(* IEC 61131-3 sources: POMIRTS_lab3/AS/Library/ETHERNET, 3 files *)

(* ---- ETHERNET.typ ---- *)
(********************************************************************
 * COPYRIGHT (C) BERNECKER + RAINER, AUSTRIA, A-5142 EGGELSBERG
 ********************************************************************
 * Library: Ethernet
 * File: Ethernet.typ
 * Created: 11.11.2003
 ********************************************************************
 * Global data types of library Ethernet
 ********************************************************************)
TYPE
	ETHattachment_typ : STRUCT
		type	: USINT ;
		len	: UDINT ;
		pName	: UDINT ;
		pData	: UDINT ;
	END_STRUCT;
	ETHstatSG3_typ : STRUCT
		l_int	: UDINT ;
		l_rint	: UDINT ;
		l_tint	: UDINT ;
		l_babl	: UINT ;
		l_cerr	: UINT ;
		l_miss	: UINT ;
		l_memr	: UINT ;
		r_fram	: UINT ;
		r_oflo	: UINT ;
		r_crc	: UINT ;
		r_buff	: UINT ;
		t_buff	: UINT ;
		t_uflo	: UINT ;
		t_lcol	: UINT ;
		t_lcar	: UINT ;
		t_rtry	: UINT ;
		ni_anno	: UINT ;
		ni_init	: UINT ;
		ni_send	: UINT ;
		ni_getp	: UINT ;
		ni_retp	: UINT ;
		ni_bcst	: UINT ;
		ni_poll	: UINT ;
		irq_mean	: UINT ;
		irq_min	: UINT ;
		irq_max	: UINT ;
		irq_t1	: UINT ;
		irq_timena	: UINT ;
		errgtnobuf	: UINT ;
		err_1_1	: UINT ;
		err_1_2	: UINT ;
		err_1_3	: UINT ;
		errxmtnull	: UINT ;
		errsndown	: UINT ;
		errsndsize	: UINT ;
		lancerrnobuf	: UINT ;
		lanceinit	: UINT ;
		terr	: UINT ;
		ni_gtbuf	: UINT ;
		brcast_cnt	: UINT ;
		brcastmax_cnt	: UINT ;
		brcast_stop	: UINT ;
		brcast_tick	: UINT ;
	END_STRUCT;
	ETHstatSG4_typ : STRUCT
		p_recv	: UDINT ;
		e_recv	: UDINT ;
		p_send	: UDINT ;
		e_send	: UDINT ;
		collisions	: UDINT ;
		b_recv	: UDINT ;
		b_send	: UDINT ;
		p_recv_mc	: UDINT ;
		p_send_mc	: UDINT ;
		iqdrops	: UDINT ;
		noproto	: UDINT ;
		lastchange	: UDINT ;
	END_STRUCT;
	TCPQ_dcmd_typ : STRUCT
		response	: UINT ;
		error	: UDINT ;
		buffer	: UDINT ;
		buflng	: UDINT ;
		ipaddr	: UDINT ;
		socket	: UDINT ;
		port	: UINT ;
		wreserve	: UINT ;
		reserve	: ARRAY[0..7] OF UDINT ;
	END_STRUCT;
END_TYPE

(* ---- ETHERNET.fun ---- *)
(********************************************************************
 * COPYRIGHT (C) BERNECKER + RAINER, AUSTRIA, A-5142 EGGELSBERG
 ********************************************************************
 * Library: Ethernet
 * File: Ethernet.fun
 * Created: 11.11.2003
 ********************************************************************
 * Functions and function blocks of library Ethernet
 ********************************************************************)
FUNCTION_BLOCK ETHinfo
	VAR_INPUT
		enable	:BOOL;
	END_VAR
	VAR_OUTPUT
		statadr	:UDINT;
		ethadr	:UDINT;
		status	:UINT;
	END_VAR
END_FUNCTION_BLOCK
FUNCTION_BLOCK SMTPxsendmail
	VAR_INPUT
		enable	:BOOL;
		pReceiver	:UDINT;
		pSender	:UDINT;
		pIpaddr	:UDINT;
		pSubject	:UDINT;
		pText	:UDINT;
		pAttachment	:UDINT;
		AttachmentCount	:USINT;
		timeout	:UINT;
	END_VAR
	VAR_OUTPUT
		status	:UINT;
	END_VAR
	VAR
		pna_ok	:BOOL;
		state	:UINT;
		tickcount	:UDINT;
		initcount	:UDINT;
		dcmd	:TCPQ_dcmd_typ;
	END_VAR
END_FUNCTION_BLOCK
FUNCTION_BLOCK ETHxinfo
	VAR_INPUT
		enable	:BOOL;
		pDevice	:UDINT;
	END_VAR
	VAR_OUTPUT
		statadr	:UDINT;
		ethadr	:UDINT;
		status	:UINT;
	END_VAR
	VAR
		mac	:ARRAY[0..5] OF USINT;
	END_VAR
END_FUNCTION_BLOCK
FUNCTION_BLOCK TCPclose
	VAR_INPUT
		enable	:BOOL;
		cident	:UDINT;
	END_VAR
	VAR_OUTPUT
		status	:UINT;
	END_VAR
	VAR
		pna_ok	:BOOL;
		state	:UINT;
		tickcount	:UDINT;
		initcount	:UDINT;
		dcmd	:TCPQ_dcmd_typ;
	END_VAR
END_FUNCTION_BLOCK
FUNCTION_BLOCK TCPrecv
	VAR_INPUT
		enable	:BOOL;
		cident	:UDINT;
		buffer	:UDINT;
		mxbuflng	:UDINT;
	END_VAR
	VAR_OUTPUT
		status	:UINT;
		rxbuflng	:UDINT;
	END_VAR
	VAR
		pna_ok	:BOOL;
		state	:UINT;
		tickcount	:UDINT;
		initcount	:UDINT;
		dcmd	:TCPQ_dcmd_typ;
	END_VAR
END_FUNCTION_BLOCK
FUNCTION_BLOCK TCPsend
	VAR_INPUT
		enable	:BOOL;
		cident	:UDINT;
		buffer	:UDINT;
		buflng	:UDINT;
	END_VAR
	VAR_OUTPUT
		status	:UINT;
	END_VAR
	VAR
		pna_ok	:BOOL;
		state	:UINT;
		tickcount	:UDINT;
		initcount	:UDINT;
		dcmd	:TCPQ_dcmd_typ;
	END_VAR
END_FUNCTION_BLOCK
FUNCTION_BLOCK TCPclient
	VAR_INPUT
		enable	:BOOL;
		porta	:UINT;
		ipaddr	:UDINT;
		portb	:UINT;
	END_VAR
	VAR_OUTPUT
		status	:UINT;
		cident	:UDINT;
	END_VAR
	VAR
		pna_ok	:BOOL;
		state	:UINT;
		tickcount	:UDINT;
		initcount	:UDINT;
		dcmd	:TCPQ_dcmd_typ;
	END_VAR
END_FUNCTION_BLOCK
FUNCTION_BLOCK TCPserv
	VAR_INPUT
		enable	:BOOL;
		porta	:UINT;
	END_VAR
	VAR_OUTPUT
		status	:UINT;
		ipaddr	:UDINT;
		portb	:UINT;
		cident	:UDINT;
	END_VAR
	VAR
		pna_ok	:BOOL;
		state	:UINT;
		tickcount	:UDINT;
		initcount	:UDINT;
		dcmd	:TCPQ_dcmd_typ;
	END_VAR
END_FUNCTION_BLOCK
FUNCTION_BLOCK ICMPping
	VAR_INPUT
		enable	:BOOL;
		ipaddr	:UDINT;
		timeout	:UINT;
	END_VAR
	VAR_OUTPUT
		status	:UINT;
	END_VAR
	VAR
		pna_ok	:BOOL;
		state	:UINT;
		tickcount	:UDINT;
		initcount	:UDINT;
		dcmd	:TCPQ_dcmd_typ;
	END_VAR
END_FUNCTION_BLOCK
FUNCTION_BLOCK SMTPsendmail
	VAR_INPUT
		enable	:BOOL;
		pReceiver	:UDINT;
		pSender	:UDINT;
		pIpaddr	:UDINT;
		pSubject	:UDINT;
		pText	:UDINT;
		timeout	:UINT;
	END_VAR
	VAR_OUTPUT
		status	:UINT;
	END_VAR
	VAR
		pna_ok	:BOOL;
		state	:UINT;
		tickcount	:UDINT;
		initcount	:UDINT;
		dcmd	:TCPQ_dcmd_typ;
	END_VAR
END_FUNCTION_BLOCK
FUNCTION_BLOCK UDPclose
	VAR_INPUT
		enable	:BOOL;
		cident	:UDINT;
	END_VAR
	VAR_OUTPUT
		status	:UINT;
	END_VAR
	VAR
		pna_ok	:BOOL;
		state	:UINT;
		tickcount	:UDINT;
		initcount	:UDINT;
		dcmd	:TCPQ_dcmd_typ;
	END_VAR
END_FUNCTION_BLOCK
FUNCTION_BLOCK UDPopen
	VAR_INPUT
		enable	:BOOL;
		port	:UINT;
		pvpolladr	:UDINT;
	END_VAR
	VAR_OUTPUT
		status	:UINT;
		cident	:UDINT;
	END_VAR
	VAR
		pna_ok	:BOOL;
		state	:UINT;
		tickcount	:UDINT;
		initcount	:UDINT;
		dcmd	:TCPQ_dcmd_typ;
	END_VAR
END_FUNCTION_BLOCK
FUNCTION_BLOCK UDPrecv
	VAR_INPUT
		enable	:BOOL;
		cident	:UDINT;
		buffer	:UDINT;
		buflng	:UINT;
	END_VAR
	VAR_OUTPUT
		status	:UINT;
		ipaddr	:UDINT;
		rxbuflng	:UINT;
		port	:UINT;
	END_VAR
	VAR
		pna_ok	:BOOL;
		state	:UINT;
		tickcount	:UDINT;
		initcount	:UDINT;
		dcmd	:TCPQ_dcmd_typ;
	END_VAR
END_FUNCTION_BLOCK
FUNCTION_BLOCK UDPsend
	VAR_INPUT
		enable	:BOOL;
		cident	:UDINT;
		ipaddr	:UDINT;
		buffer	:UDINT;
		buflng	:UINT;
		port	:UINT;
	END_VAR
	VAR_OUTPUT
		status	:UINT;
	END_VAR
	VAR
		pna_ok	:BOOL;
		state	:UINT;
		tickcount	:UDINT;
		initcount	:UDINT;
		dcmd	:TCPQ_dcmd_typ;
	END_VAR
END_FUNCTION_BLOCK
FUNCTION_BLOCK ETHnode
	VAR_INPUT
		enable	:BOOL;
	END_VAR
	VAR_OUTPUT
		status	:UINT;
		nodenr	:USINT;
		ipaddr	:UDINT;
	END_VAR
	VAR
		address1	:UDINT;
		address2	:UDINT;
	END_VAR
END_FUNCTION_BLOCK

(* ---- ETHERNET.var ---- *)
(********************************************************************
 * COPYRIGHT (C) BERNECKER + RAINER, AUSTRIA, A-5142 EGGELSBERG
 ********************************************************************
 * Library: Ethernet
 * File: Ethernet.var
 * Created: 11.11.2003
 ********************************************************************
 * Constants of library Ethernet
 ********************************************************************)
VAR CONSTANT
	ERR_ETH_SMTP_UNEXPECTED_RESPONSE	: UINT	:= 27232;
	ERR_ETH_SMTP_SERVER_NOTAVAILABLE	: UINT	:= 27230;
	ERR_ETH_SMTP_RECEIVER_NOT_ACCEPT	: UINT	:= 27234;
	ERR_ETH_SMTP_PARSE_NO_SEMI_COLON	: UINT	:= 27233;
	ERR_ETH_SMTP_MAIL_CANNOT_DELIVER	: UINT	:= 27235;
	ERR_ETH_INVALID_ATTACHMENT	: UINT	:= 27240;
	ERR_ETH_SMTP_TIMEOUT	: UINT	:= 27231;
	ERR_ETH_PING_TIMEOUT	: UINT	:= 27221;
	ERR_ETH_DEVICE_ERROR	: UINT	:= 27247;
	ERR_ETH_PING_NORESP	: UINT	:= 27220;
	ETH_ATT_TYPE_FILE	: USINT	:= 1;
	ETH_ATT_TYPE_MEM	: USINT	:= 0;
	ERR_ETH_NET_SLOW	: UINT	:= 27210;
	ERR_ETH_NO_DATA	: UINT	:= 27211;
END_VAR
